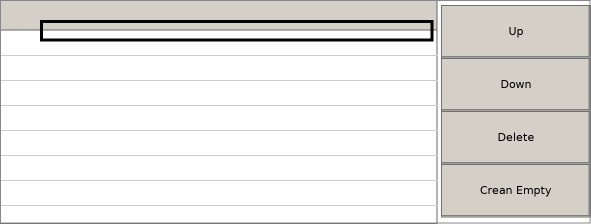
VISUALIZATION vis_CIP_ReqBuffer  // 591x224
    Table (0,0 437x224), data array: arCIP_RequestBufer
        p1137915858: fbCIP.iPosSelect_HMI
        p3854506369: arCIP_RequestBufer[INDEX].eType
        p1892666644: arCIP_RequestBufer[INDEX].eClient
    Button (441,5 150x53), "Up"
        tap fbCIP.rtPosMoveHMI_Up.CLK
    Button (441,58 150x53), "Down"
        tap fbCIP.rtPosMoveHMI_Down.CLK
    Button (441,111 150x53), "Delete"
        tap fbCIP.rtPosDeleteHMI.CLK
    Rectangle (40,20 393x21), colour toggle: fbCIP.bRun
    Button (441,164 150x53), "Crean Empty"
        tap fbCIP.rtReqCleanEmpty_HMI.CLK
END_VISUALIZATION

(* stored: Version 1.1.0.1, ProductVersion 3.1.4024.12
   Visu vis_CIP_ReqBuffer: Id {5967227b-2f86-4543-bece-239394dbe74e} *)
